// SIMATIC S7-200 project (STEP 7-Micro/WIN), CPU 226 CN REL 02.01

SYMBOL_TABLE 用户定义1
允许装配             V1000.5
停止               M0.1
准备就绪             M0.0
缺料               V1010.3
料不足              V1010.2
全线模式             V1010.1
网络正常             V1010.0
装配完成             V1010.4
急停               V1010.5
故障无法修复           V1010.6
物料不足检测           I0.0
物料有无检测           I0.1
物料左检测            I0.2
物料右检测            I0.3
物料台检测            I0.4
顶料到位检测           I0.5
顶料复位检测           I0.6
挡料状态检测           I0.7
落料状态检测           I1.0
旋转缸左限位检测         I1.1
旋转缸右限位检测         I1.2
手抓夹紧检测           I1.3
手抓下降到位检测         I1.4
手抓上升到位检测         I1.5
手抓缩回到位检测         I1.6
手抓伸出到位检测         I1.7
停止按钮             I2.4
启动按钮             I2.5
急停按钮             I2.6
单机全线             I2.7
挡料电磁阀            Q0.0
顶料电磁阀            Q0.1
回转电磁阀            Q0.2
手抓夹紧电磁阀          Q0.3
手抓下降电磁阀          Q0.4     // .
手抓伸出电磁阀          Q0.5
红色警示灯            Q0.6
黄色警示灯            Q0.7
绿色警示灯            Q1.0
黄色指示灯            Q1.5
绿色指示灯            Q1.6
红色指示灯            Q1.7
END_SYMBOL_TABLE

ORGANIZATION_BLOCK 主程序:OB1
TITLE=程序注释
BEGIN
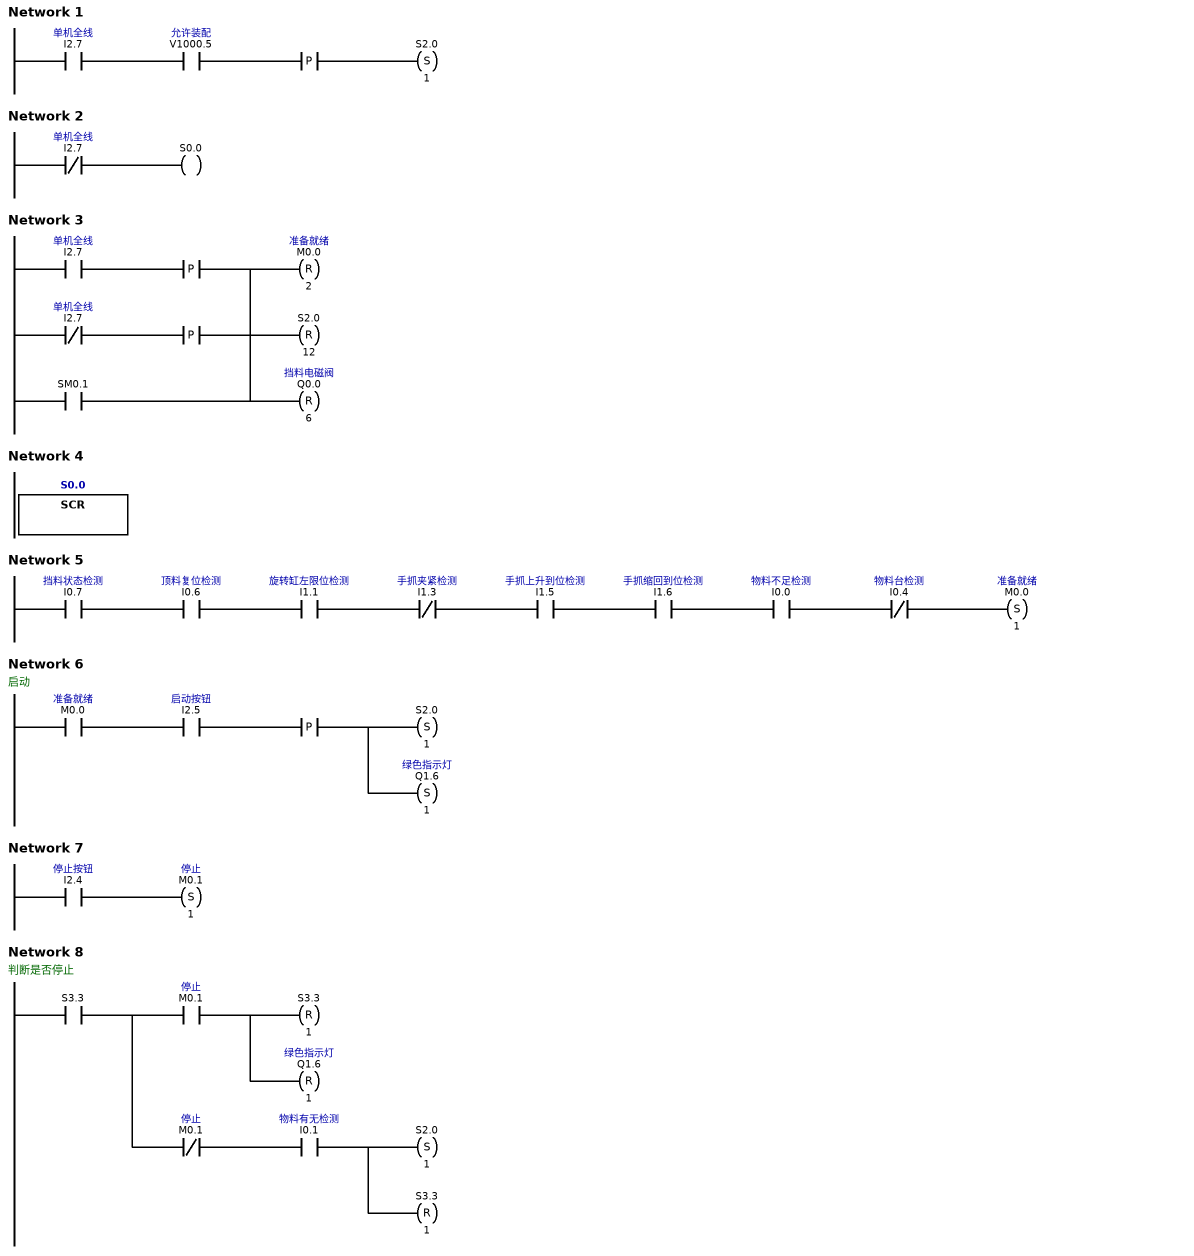
Network 1
LD     单机全线:I2.7
A      允许装配:V1000.5
EU
S      S2.0, 1
Network 2
LDN    单机全线:I2.7
=      S0.0
Network 3
LD     单机全线:I2.7
EU
LDN    单机全线:I2.7
EU
OLD
O      SM0.1
R      准备就绪:M0.0, 2
R      S2.0, 12
R      挡料电磁阀:Q0.0, 6
Network 4
LSCR   S0.0
Network 5
LD     挡料状态检测:I0.7
A      顶料复位检测:I0.6
A      旋转缸左限位检测:I1.1
AN     手抓夹紧检测:I1.3
A      手抓上升到位检测:I1.5
A      手抓缩回到位检测:I1.6
A      物料不足检测:I0.0
AN     物料台检测:I0.4
S      准备就绪:M0.0, 1
Network 6
// 启动
LD     准备就绪:M0.0
A      启动按钮:I2.5
EU
S      S2.0, 1
S      绿色指示灯:Q1.6, 1
Network 7
LD     停止按钮:I2.4
S      停止:M0.1, 1
Network 8
// 判断是否停止
LD     S3.3
LPS
A      停止:M0.1
R      S3.3, 1
R      绿色指示灯:Q1.6, 1
LPP
AN     停止:M0.1
A      物料有无检测:I0.1
S      S2.0, 1
R      S3.3, 1
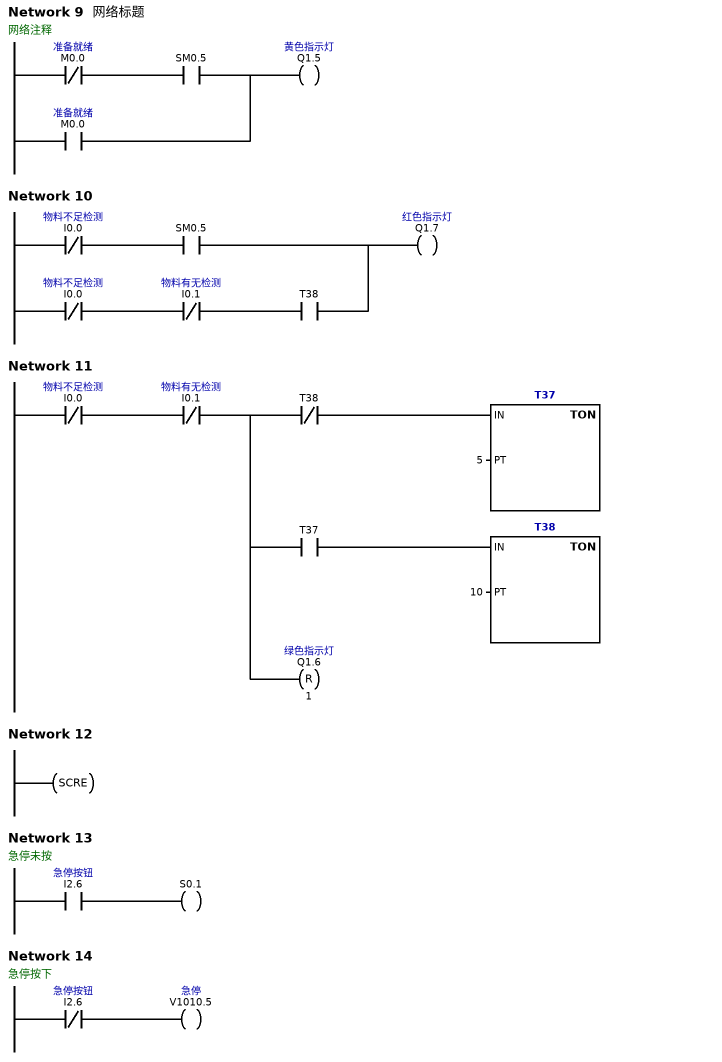
Network 9 // 网络标题
// 网络注释
LDN    准备就绪:M0.0
A      SM0.5
O      准备就绪:M0.0
=      黄色指示灯:Q1.5
Network 10
LDN    物料不足检测:I0.0
A      SM0.5
LDN    物料不足检测:I0.0
AN     物料有无检测:I0.1
A      T38
OLD
=      红色指示灯:Q1.7
Network 11
LDN    物料不足检测:I0.0
AN     物料有无检测:I0.1
LPS
AN     T38
TON    T37, 5
LRD
A      T37
TON    T38, 10
LPP
R      绿色指示灯:Q1.6, 1
Network 12
SCRE
Network 13
// 急停未按
LD     急停按钮:I2.6
=      S0.1
Network 14
// 急停按下
LDN    急停按钮:I2.6
=      急停:V1010.5
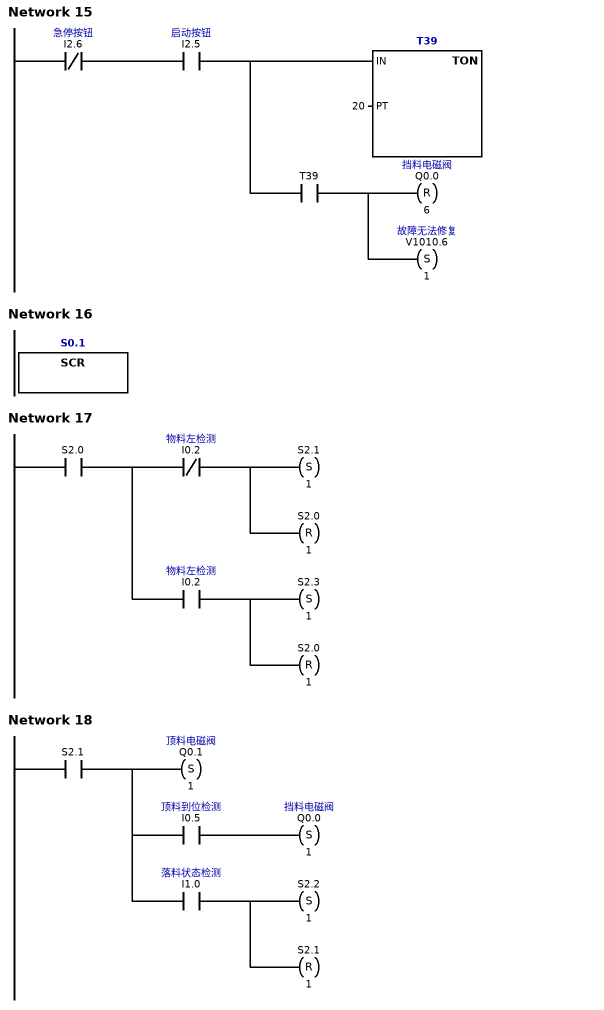
Network 15
LDN    急停按钮:I2.6
A      启动按钮:I2.5
TON    T39, 20
A      T39
R      挡料电磁阀:Q0.0, 6
S      故障无法修复:V1010.6, 1
Network 16
LSCR   S0.1
Network 17
LD     S2.0
LPS
AN     物料左检测:I0.2
S      S2.1, 1
R      S2.0, 1
LPP
A      物料左检测:I0.2
S      S2.3, 1
R      S2.0, 1
Network 18
LD     S2.1
LPS
S      顶料电磁阀:Q0.1, 1
A      顶料到位检测:I0.5
S      挡料电磁阀:Q0.0, 1
LPP
A      落料状态检测:I1.0
S      S2.2, 1
R      S2.1, 1
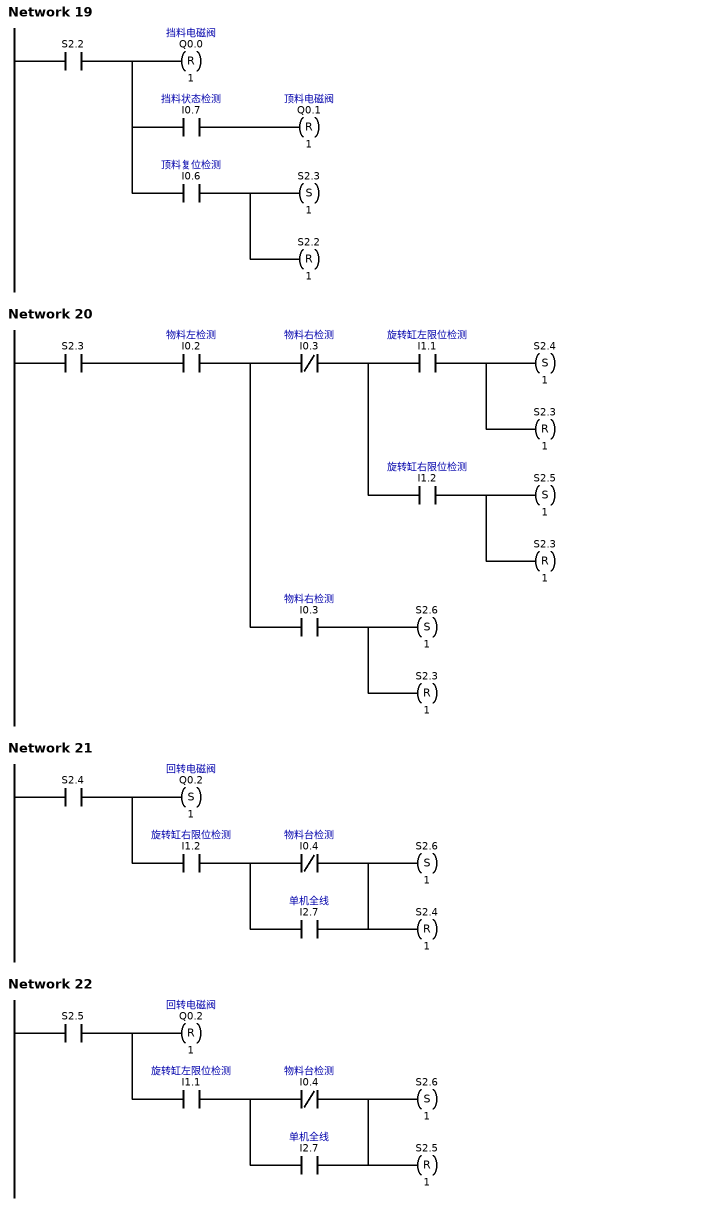
Network 19
LD     S2.2
LPS
R      挡料电磁阀:Q0.0, 1
A      挡料状态检测:I0.7
R      顶料电磁阀:Q0.1, 1
LPP
A      顶料复位检测:I0.6
S      S2.3, 1
R      S2.2, 1
Network 20
LD     S2.3
A      物料左检测:I0.2
LPS
AN     物料右检测:I0.3
LPS
A      旋转缸左限位检测:I1.1
S      S2.4, 1
R      S2.3, 1
LPP
A      旋转缸右限位检测:I1.2
S      S2.5, 1
R      S2.3, 1
LPP
A      物料右检测:I0.3
S      S2.6, 1
R      S2.3, 1
Network 21
LD     S2.4
S      回转电磁阀:Q0.2, 1
A      旋转缸右限位检测:I1.2
LDN    物料台检测:I0.4
O      单机全线:I2.7
ALD
S      S2.6, 1
R      S2.4, 1
Network 22
LD     S2.5
R      回转电磁阀:Q0.2, 1
A      旋转缸左限位检测:I1.1
LDN    物料台检测:I0.4
O      单机全线:I2.7
ALD
S      S2.6, 1
R      S2.5, 1
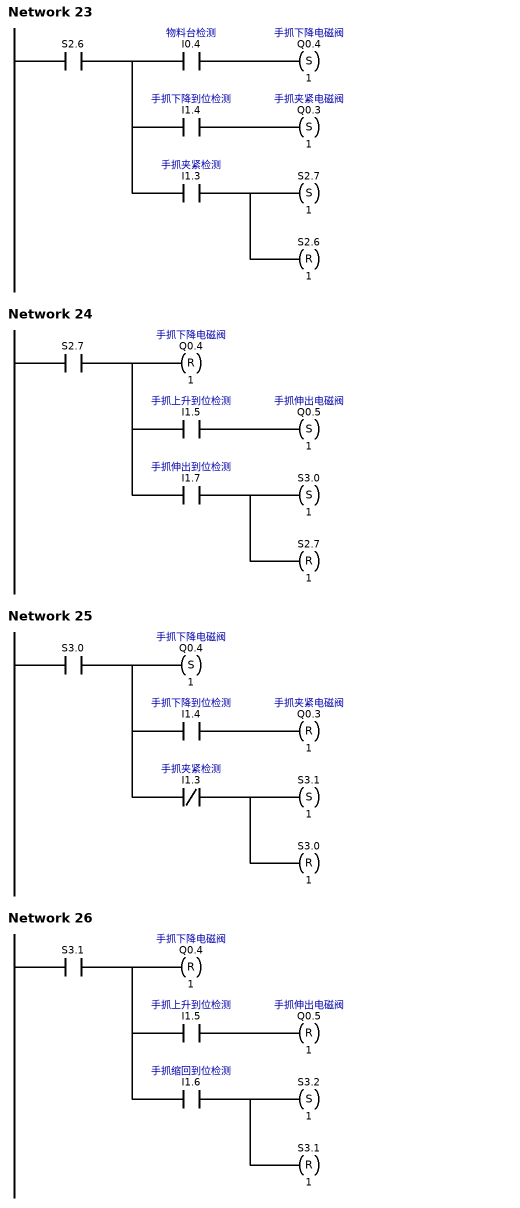
Network 23
LD     S2.6
LPS
A      物料台检测:I0.4
S      手抓下降电磁阀:Q0.4, 1
LRD
A      手抓下降到位检测:I1.4
S      手抓夹紧电磁阀:Q0.3, 1
LPP
A      手抓夹紧检测:I1.3
S      S2.7, 1
R      S2.6, 1
Network 24
LD     S2.7
LPS
R      手抓下降电磁阀:Q0.4, 1
A      手抓上升到位检测:I1.5
S      手抓伸出电磁阀:Q0.5, 1
LPP
A      手抓伸出到位检测:I1.7
S      S3.0, 1
R      S2.7, 1
Network 25
LD     S3.0
LPS
S      手抓下降电磁阀:Q0.4, 1
A      手抓下降到位检测:I1.4
R      手抓夹紧电磁阀:Q0.3, 1
LPP
AN     手抓夹紧检测:I1.3
S      S3.1, 1
R      S3.0, 1
Network 26
LD     S3.1
LPS
R      手抓下降电磁阀:Q0.4, 1
A      手抓上升到位检测:I1.5
R      手抓伸出电磁阀:Q0.5, 1
LPP
A      手抓缩回到位检测:I1.6
S      S3.2, 1
R      S3.1, 1
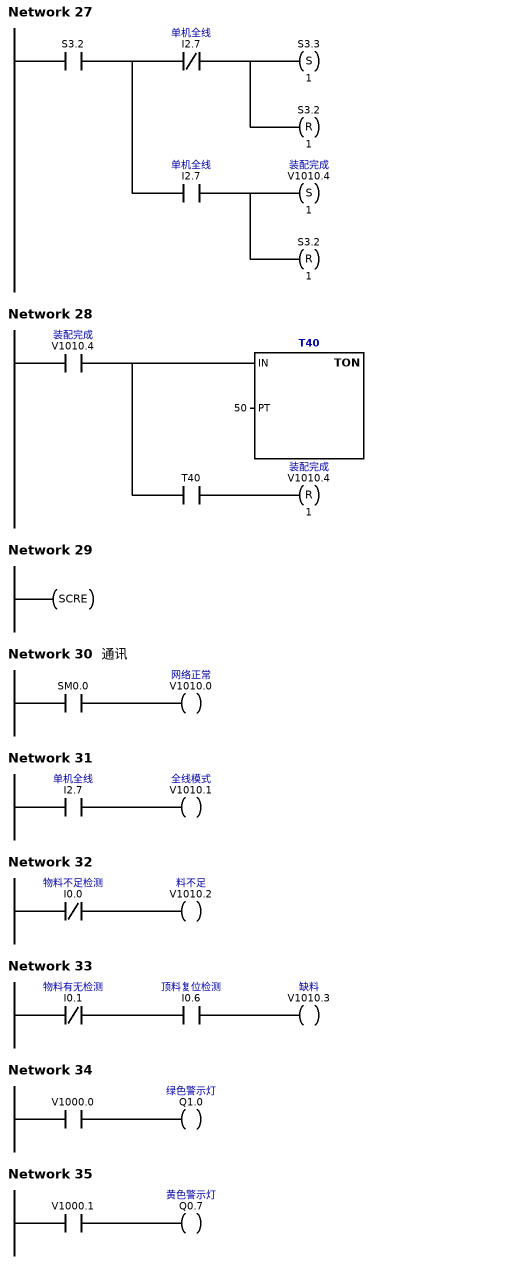
Network 27
LD     S3.2
LPS
AN     单机全线:I2.7
S      S3.3, 1
R      S3.2, 1
LPP
A      单机全线:I2.7
S      装配完成:V1010.4, 1
R      S3.2, 1
Network 28
LD     装配完成:V1010.4
TON    T40, 50
A      T40
R      装配完成:V1010.4, 1
Network 29
SCRE
Network 30 // 通讯
LD     SM0.0
=      网络正常:V1010.0
Network 31
LD     单机全线:I2.7
=      全线模式:V1010.1
Network 32
LDN    物料不足检测:I0.0
=      料不足:V1010.2
Network 33
LDN    物料有无检测:I0.1
A      顶料复位检测:I0.6
=      缺料:V1010.3
Network 34
LD     V1000.0
=      绿色警示灯:Q1.0
Network 35
LD     V1000.1
=      黄色警示灯:Q0.7
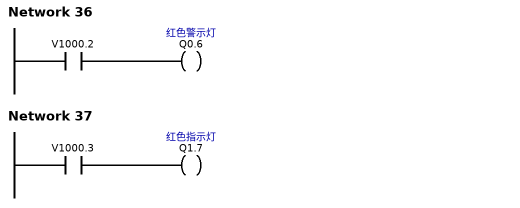
Network 36
LD     V1000.2
=      红色警示灯:Q0.6
Network 37
LD     V1000.3
=      红色指示灯:Q1.7
END_ORGANIZATION_BLOCK
